Fanuc KAREL source: kt00130.KL

-- PROVISIONAL review KL for V940-1; original PC SHA256 c5cc95534a2d6f8d86ac34434cd2ded4dd8563663df0d4bc0c7240e95a850335
-- Incomplete behavior may be omitted. Consult companion uncertainty JSON. Do not deploy.
PROGRAM KT00130
%NOLOCKGROUP
VAR
  I1 : INTEGER
  I2 : INTEGER
  OUT : REAL
BEGIN
  -- V9_ZERO_TABLE_METADATA_HINT layout=0001; no indexed target words; source/name/runtime held
  -- UNRESOLVED_PC offsets 5-16; opcodes 2E,23
  -- UNRESOLVED_PC offsets 21-32; opcodes 2E,23
  -- UNRESOLVED_PC offsets 37-48; opcodes 2E,23
  -- UNRESOLVED_PC offsets 53-64; opcodes 2E,23
  -- UNRESOLVED_PC offsets 69-89; opcodes 21,21,55,64,23
  -- UNRESOLVED_PC offsets 94-98; opcodes 7F
END KT00130
